(* IEC 61131-3 sources: trust-platform/examples/control/01-feedback-foundations-and-temperature-control/17-gravity-tank-linearization/src, 2 files *)

(* ---- Main.st ---- *)
(* Slope of the gravity outflow q = c·√h at the operating level h0: g = c/(2·√h0), in m²/s. *)
FUNCTION TangentSlope : LREAL
VAR_INPUT
    Coefficient : LREAL;
    OperatingLevel : LREAL;
END_VAR
TangentSlope := Coefficient / (LREAL#2.0 * SQRT(OperatingLevel));
END_FUNCTION

(* One update of the tangent model A·dx/dt = v − g·x, for the level deviation x and the inflow deviation v. *)
FUNCTION TangentDeviationNext : LREAL
VAR_INPUT
    Deviation : LREAL;
    InflowDeviation : LREAL;
    Slope : LREAL;
    Area : LREAL;
    CycleTime : LREAL;
END_VAR
TangentDeviationNext := Deviation + (InflowDeviation - Slope * Deviation) / Area * CycleTime;
END_FUNCTION

PROGRAM Main
VAR
    (* Two identical tanks of Lesson 45 (A = 0.5 m², c = 0.020 m^(5/2)/s), both operating at h0 = 0.25 m with
       q0 = 0.010 m³/s. *)
    TankAreaM2 : LREAL := 0.5;
    OutletCoefficient : LREAL := 0.020;
    OperatingLevelM : LREAL := 0.25;
    OperatingFlowM3S : LREAL := 0.010;
    TangentSlopeM2S : LREAL := 0.0;
    SmallInletFlowM3S : LREAL := 0.010;
    LargeInletFlowM3S : LREAL := 0.010;
    (* The measured levels, in m. The program only reads them. *)
    SmallLevelM : LREAL := 0.0;
    LargeLevelM : LREAL := 0.0;
    (* The tangent models: deviations from h0, advanced every 1 s update with the inflow deviation applied during
       that second and started from the measured levels. *)
    SmallDeviationM : LREAL := 0.0;
    LargeDeviationM : LREAL := 0.0;
    SmallTangentLevelM : LREAL := 0.0;
    LargeTangentLevelM : LREAL := 0.0;
    AppliedSmallInletM3S : LREAL := 0.010;
    AppliedLargeInletM3S : LREAL := 0.010;
    ModelStarted : BOOL := FALSE;
    (* Control Studio's project experiment: 0.011 m³/s into one tank and 0.015 m³/s into the other while it runs. *)
    ExperimentEnabled : BOOL := FALSE;
    ExperimentWasEnabled : BOOL := FALSE;
    Active : BOOL := FALSE;
END_VAR

TangentSlopeM2S := TangentSlope(Coefficient := OutletCoefficient, OperatingLevel := OperatingLevelM);
IF NOT ModelStarted THEN
    SmallDeviationM := SmallLevelM - OperatingLevelM;
    LargeDeviationM := LargeLevelM - OperatingLevelM;
    ModelStarted := TRUE;
ELSE
    SmallDeviationM := TangentDeviationNext(Deviation := SmallDeviationM, InflowDeviation := AppliedSmallInletM3S - OperatingFlowM3S,
        Slope := TangentSlopeM2S, Area := TankAreaM2, CycleTime := LREAL#1.0);
    LargeDeviationM := TangentDeviationNext(Deviation := LargeDeviationM, InflowDeviation := AppliedLargeInletM3S - OperatingFlowM3S,
        Slope := TangentSlopeM2S, Area := TankAreaM2, CycleTime := LREAL#1.0);
END_IF;

IF ExperimentEnabled AND NOT ExperimentWasEnabled THEN
    Active := TRUE;
    (* Each experiment compares from the levels measured at its step. *)
    SmallDeviationM := SmallLevelM - OperatingLevelM;
    LargeDeviationM := LargeLevelM - OperatingLevelM;
ELSIF NOT ExperimentEnabled THEN
    Active := FALSE;
END_IF;
ExperimentWasEnabled := ExperimentEnabled;
SmallTangentLevelM := OperatingLevelM + SmallDeviationM;
LargeTangentLevelM := OperatingLevelM + LargeDeviationM;

IF Active THEN
    SmallInletFlowM3S := LREAL#0.011;
    LargeInletFlowM3S := LREAL#0.015;
ELSE
    SmallInletFlowM3S := LREAL#0.010;
    LargeInletFlowM3S := LREAL#0.010;
END_IF;
AppliedSmallInletM3S := SmallInletFlowM3S;
AppliedLargeInletM3S := LargeInletFlowM3S;
END_PROGRAM

CONFIGURATION Config
RESOURCE Res ON PLC
    TASK MainTask(INTERVAL := T#1s, PRIORITY := 1);
    PROGRAM P1 WITH MainTask : Main;
END_RESOURCE
VAR_CONFIG
    P1.SmallInletFlowM3S AT %QL0 : LREAL;
    P1.LargeInletFlowM3S AT %QL8 : LREAL;
    P1.SmallLevelM AT %IL0 : LREAL;
    P1.LargeLevelM AT %IL8 : LREAL;
    P1.SmallTangentLevelM AT %ML0 : LREAL;
    P1.LargeTangentLevelM AT %ML8 : LREAL;
    P1.ExperimentEnabled AT %MX16.0 : BOOL;
    P1.Active AT %MX16.1 : BOOL;
END_VAR
END_CONFIGURATION

(* ---- tests.st ---- *)
(* @trustlsp:runtime-ignore — run these assertions with trust-dev test;
   they are not scheduled PLC instances in the lesson simulator. *)

TEST_PROGRAM TheTangentAtTheOperatingLevel
VAR
    Slope : LREAL;
END_VAR
(* c = 0.020 m^(5/2)/s at h0 = 0.25 m: g = 0.020/(2 · 0.5) = 0.020 m²/s, K = 1/g = 50 s/m², τ = A/g = 25 s. *)
Slope := TangentSlope(Coefficient := LREAL#0.020, OperatingLevel := LREAL#0.25);
ASSERT_NEAR(EXPECTED := LREAL#0.020, ACTUAL := Slope, DELTA := LREAL#1.0e-12);
ASSERT_NEAR(EXPECTED := LREAL#50.0, ACTUAL := LREAL#1.0 / Slope, DELTA := LREAL#1.0e-9);
ASSERT_NEAR(EXPECTED := LREAL#25.0, ACTUAL := LREAL#0.5 / Slope, DELTA := LREAL#1.0e-9);
END_TEST_PROGRAM

TEST_PROGRAM TheTangentErrorGrowsWithTheSquareOfTheStep
(* Tangent equilibria h0 + v/g: 0.3000 m for v = 0.001 and 0.5000 m for v = 0.005 m³/s. Exact equilibria
   (q/c)²: 0.3025 m and 0.5625 m. The difference is v²/c²: 0.0025 m and 0.0625 m, 25 times more for 5 times
   the step. A 0.005 m error allows |v| ≤ c·√0.005 = 0.00141 m³/s. *)
ASSERT_NEAR(EXPECTED := LREAL#0.3000, ACTUAL := LREAL#0.25 + LREAL#0.001 / LREAL#0.020, DELTA := LREAL#1.0e-12);
ASSERT_NEAR(EXPECTED := LREAL#0.5000, ACTUAL := LREAL#0.25 + LREAL#0.005 / LREAL#0.020, DELTA := LREAL#1.0e-12);
ASSERT_NEAR(EXPECTED := LREAL#0.3025 - LREAL#0.3000, ACTUAL := (LREAL#0.001 / LREAL#0.020) * (LREAL#0.001 / LREAL#0.020),
    DELTA := LREAL#1.0e-12);
ASSERT_NEAR(EXPECTED := LREAL#0.5625 - LREAL#0.5000, ACTUAL := (LREAL#0.005 / LREAL#0.020) * (LREAL#0.005 / LREAL#0.020),
    DELTA := LREAL#1.0e-12);
ASSERT_NEAR(EXPECTED := LREAL#0.001414, ACTUAL := LREAL#0.020 * SQRT(LREAL#0.005), DELTA := LREAL#1.0e-6);
END_TEST_PROGRAM
